FUNCTION_BLOCK AOption_OR_3 (* Options-Fan-In: 3 AOption-Sockets IN1/IN2/IN3 auf 1 Plug OUT, QI_OUT = IN1 ODER IN2 ODER IN3. OUT.INIT_CNF geht per E_MUX_3/E_DEMUX_3 an den anfragenden Socket zurueck. *)
  (* Standard: 61499-1; Description: Copyright (c) 2026 Meisterschulen am Ostbahnhof This program and the accompanying materials are made available under the terms of the Eclipse Public License 2.0 which is available at https://www.eclipse.org/legal/epl-2.0/ SPDX-License-Identifier: EPL-2.0 *)
  (* Version 1.0, 2026-10-17, Franz Höpfinger, Meisterschulen am Ostbahnhof, Wie AOption_OR_2 mit 3 Eingaengen. E_MUX_3.K merkt den anfragenden Socket, E_DEMUX_3 leitet OUT.INIT_CNF dorthin. Max. 1 offene Anfrage. *)
  PACKAGE Option::merging;
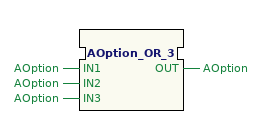
  SOCKETS
    IN1 : Option::AOption; (* Erster AOption-Eingang *)
    IN2 : Option::AOption; (* Zweiter AOption-Eingang *)
    IN3 : Option::AOption; (* Dritter AOption-Eingang *)
  END_SOCKETS
  PLUGS
    OUT : Option::AOption; (* Gemeinsamer Ausgang - aktiv, solange IN1 ODER IN2 ODER IN3 aktiv ist *)
  END_PLUGS
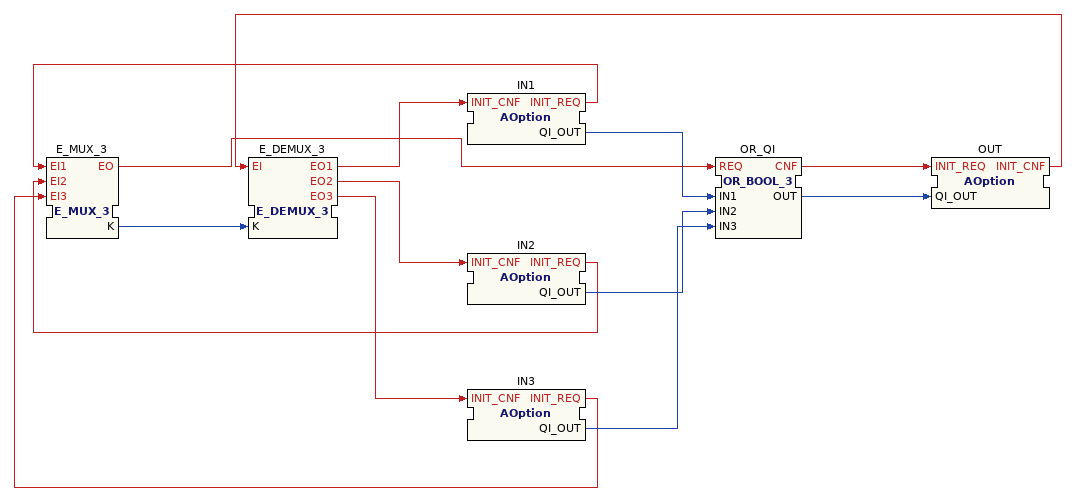
  FBS
    OR_QI : iec61131::booleanOperators::OR_BOOL_3;
    E_MUX_3 : iec61499::events::E_MUX_3;
    E_DEMUX_3 : iec61499::events::E_DEMUX_3;
  END_FBS
  EVENT_CONNECTIONS
    OR_QI.CNF TO OUT.INIT_REQ;
    OUT.INIT_CNF TO E_DEMUX_3.EI;
    E_DEMUX_3.EO1 TO IN1.INIT_CNF;
    E_DEMUX_3.EO2 TO IN2.INIT_CNF;
    E_DEMUX_3.EO3 TO IN3.INIT_CNF;
    IN1.INIT_REQ TO E_MUX_3.EI1;
    IN2.INIT_REQ TO E_MUX_3.EI2;
    IN3.INIT_REQ TO E_MUX_3.EI3;
    E_MUX_3.EO TO OR_QI.REQ;
  END_CONNECTIONS
  DATA_CONNECTIONS
    IN1.QI_OUT TO OR_QI.IN1;
    IN2.QI_OUT TO OR_QI.IN2;
    IN3.QI_OUT TO OR_QI.IN3;
    OR_QI.OUT TO OUT.QI_OUT;
    E_MUX_3.K TO E_DEMUX_3.K;
  END_CONNECTIONS
END_FUNCTION_BLOCK
